FUNCTION_BLOCK Desinfeccao_UV_HMI (* Service Interface Function Block Type *)
  (* Standard: 61499-2 *)
  (* Version 1.1, 21/10/2026, Hidryco, Hidryco, IHM da Desinfeccao_UV 1.1: ajustes do PID no sub-CAT PID_VC_700_01; reset cmdResetFalhas / E_RESET_FALHAS_PROCESSO (legado) *)
  PACKAGE Hidryco.HidrycoLib;
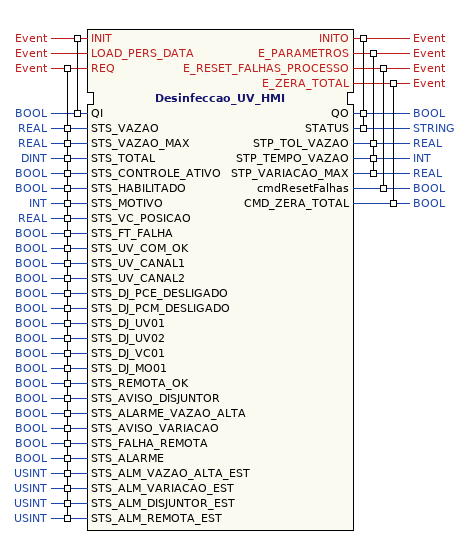
  EVENT_INPUT
    INIT WITH QI;
    LOAD_PERS_DATA; (* Reenvia os parametros persistentes *)
    REQ WITH STS_VAZAO, STS_VAZAO_MAX, STS_TOTAL, STS_CONTROLE_ATIVO, STS_HABILITADO, STS_MOTIVO, STS_VC_POSICAO, STS_FT_FALHA, STS_UV_COM_OK, STS_UV_CANAL1, STS_UV_CANAL2, STS_DJ_PCE_DESLIGADO, STS_DJ_PCM_DESLIGADO, STS_DJ_UV01, STS_DJ_UV02, STS_DJ_VC01, STS_DJ_MO01, STS_REMOTA_OK, STS_AVISO_DISJUNTOR, STS_ALARME_VAZAO_ALTA, STS_AVISO_VARIACAO, STS_FALHA_REMOTA, STS_ALARME, STS_ALM_VAZAO_ALTA_EST, STS_ALM_VARIACAO_EST, STS_ALM_DISJUNTOR_EST, STS_ALM_REMOTA_EST; (* Atualizacao de status *)
  END_EVENT
  EVENT_OUTPUT
    INITO WITH QO, STATUS;
    E_PARAMETROS WITH STP_TOL_VAZAO, STP_TEMPO_VAZAO, STP_VARIACAO_MAX;
    E_RESET_FALHAS_PROCESSO WITH cmdResetFalhas;
    E_ZERA_TOTAL WITH CMD_ZERA_TOTAL;
  END_EVENT
  VAR_INPUT
    QI : BOOL;
    STS_VAZAO : REAL; (* Vazao do efluente final 700-FT-01 (m3/h) *)
    STS_VAZAO_MAX : REAL; (* Vazao maxima de lancamento em uso (m3/h) *)
    STS_TOTAL : DINT; (* Volume totalizado (m3) *)
    STS_CONTROLE_ATIVO : BOOL; (* PID controlando a 700-VC-01 *)
    STS_HABILITADO : BOOL; (* Controle de vazao habilitado pelo operador *)
    STS_MOTIVO : INT; (* Controle: 0 controlando, 1 desabilitado, 2 FT-01 em falha, 3 valvula indisponivel, 4 retomando (3 s) *)
    STS_VC_POSICAO : REAL; (* Posicao da 700-VC-01 (%) *)
    STS_FT_FALHA : BOOL; (* 700-FT-01 em falha *)
    STS_UV_COM_OK : BOOL; (* UV comunicando *)
    STS_UV_CANAL1 : BOOL; (* UV canal 1 operando *)
    STS_UV_CANAL2 : BOOL; (* UV canal 2 operando *)
    STS_DJ_PCE_DESLIGADO : BOOL; (* Remota %I0.0: disjuntor desligado PCE *)
    STS_DJ_PCM_DESLIGADO : BOOL; (* Remota %I0.1: disjuntor desligado PCM desinfeccao *)
    STS_DJ_UV01 : BOOL; (* Remota %I0.2: disjuntor ligado 700-UV-01 *)
    STS_DJ_UV02 : BOOL; (* Remota %I0.3: disjuntor ligado 700-UV-02 *)
    STS_DJ_VC01 : BOOL; (* Remota %I0.4: disjuntor ligado 700-VC-01 *)
    STS_DJ_MO01 : BOOL; (* Remota %I0.5: disjuntor ligado 700-MO-01 (monovia) *)
    STS_REMOTA_OK : BOOL; (* Remota da desinfeccao comunicando *)
    STS_AVISO_DISJUNTOR : BOOL; (* Disjuntor do PCE, PCM, UV ou VC-01 desligado *)
    STS_ALARME_VAZAO_ALTA : BOOL; (* Vazao acima do limite de lancamento (memorizado) *)
    STS_AVISO_VARIACAO : BOOL; (* Variacao brusca da vazao de lancamento (memorizado) *)
    STS_FALHA_REMOTA : BOOL; (* Falha de comunicacao com a remota da desinfeccao *)
    STS_ALARME : BOOL; (* Algum alarme da desinfeccao *)
    STS_ALM_VAZAO_ALTA_EST : USINT; (* Estado do ALARM_BIT (0 normal, 1 ativo reconhecido, 2 ativo nao reconhecido, 3 saiu nao reconhecido, 4 ativo e saiu nao reconhecido) *)
    STS_ALM_VARIACAO_EST : USINT; (* Estado do ALARM_BIT (0 normal, 1 ativo reconhecido, 2 ativo nao reconhecido, 3 saiu nao reconhecido, 4 ativo e saiu nao reconhecido) *)
    STS_ALM_DISJUNTOR_EST : USINT; (* Estado do ALARM_BIT (0 normal, 1 ativo reconhecido, 2 ativo nao reconhecido, 3 saiu nao reconhecido, 4 ativo e saiu nao reconhecido) *)
    STS_ALM_REMOTA_EST : USINT; (* Estado do ALARM_BIT (0 normal, 1 ativo reconhecido, 2 ativo nao reconhecido, 3 saiu nao reconhecido, 4 ativo e saiu nao reconhecido) *)
  END_VAR
  VAR_OUTPUT
    QO : BOOL; (* Event Output Qualifier *)
    STATUS : STRING; (* Service Status *)
    STP_TOL_VAZAO : REAL; (* Alarme: tolerancia acima do limite (%) *)
    STP_TEMPO_VAZAO : INT; (* Alarme: tempo acima do limite (s); 0 = desligado *)
    STP_VARIACAO_MAX : REAL; (* Aviso: variacao maxima da vazao em 1 min (m3/h); 0 = desligado *)
    cmdResetFalhas : BOOL; (* Reconhece os alarmes da desinfeccao *)
    CMD_ZERA_TOTAL : BOOL; (* Zera o totalizador *)
  END_VAR
  SERVICE /
    SEQUENCE 
    END_SEQUENCE
  END_SERVICE
END_FUNCTION_BLOCK
